{attribute 'Tc2GvlVarNames'}
VAR_GLOBAL CONSTANT
	usnFileArrayMaxDimR					:USINT := 100;		(* 0..usnMaxDimR - Number of rows to read. *)
	usnFileArrayMaxDimC					:USINT := 1;  			(* 0..usnMaxDimC -  Number of columns to read. *)
END_VAR

(* stored: Version 1.1.0.1, ProductVersion 3.1.4024.15
   GVL GVL_FB_LoadFromFile: Id {83c15935-6d48-40d3-b6da-0535fcab9b8d} *)
